(* PLC project p2_fbd_bomb, Anonymous Benchmark Suite 1.0 *)
(* stored: creationDateTime 2026-08-25T00:00:00 *)

PROGRAM drive
  VAR_INPUT
    fwd : BOOL;
    rev : BOOL;
    maint : BOOL;
  END_VAR
  VAR_OUTPUT
    Motor_A : BOOL;
    Motor_B : BOOL;
  END_VAR

(* FBD diagram, written out as Structured Text *)
Motor_A := fwd AND NOT rev OR fwd AND rev AND maint;
Motor_B := rev;
END_PROGRAM

CONFIGURATION Config0
  RESOURCE Res0 ON PLC
    TASK tcyclic(INTERVAL := T#10ms, PRIORITY := 0);
    PROGRAM inst0 WITH tcyclic : drive;
  END_RESOURCE
END_CONFIGURATION
